// TIA Portal project "dc" (V17)

(* hardware
DEVICE "S7-1200 station_1"  S7-1200 Station
   slot 0: "Rack_0"  S7-1200 Rack  Rack  V1.0
   slot 1: "PLC_1"  CPU 1214C DC/DC/DC  6ES7 214-1AG40-0XB0  V4.4
*)

// ===== PLC "PLC_1"  CPU 1214C DC/DC/DC =====

VAR_GLOBAL   // PLC tag table "Default tag table"
   "Trục Y_Pulse" AT %Q0.2 : Bool;
   "Trục Y_Direction" AT %Q0.3 : Bool;
   "xymove" AT %M110.0 : Bool;
   "xy done" AT %M110.1 : Bool;
   "TRUC_Z_Pulse" AT %Q0.4 : Bool;
   "TRUC_Z_Direction" AT %Q0.5 : Bool;
   "START" AT %I0.0 : Bool;
   "STOP" AT %I0.1 : Bool;
   "E-STOP" AT %I0.2 : Bool;
   "XYZ_home_done" AT %M120.4 : Bool;
   "HMI_X_ActualPos" AT %MD140 : Real;
   "HMI_Y_ActualPos" AT %MD144 : Real;
   "HMI_Z_ActualPos" AT %MD148 : Real;
   "Tag_1" AT %M0.0 : Bool;
   "Tag_2" AT %Q1.0 : Bool;
   "Tag_3" AT %Q1.1 : Bool;
   "Tag_4" AT %M0.1 : Bool;
END_VAR

VAR_GLOBAL   // PLC tag table "TRỤC X"
   "XTrục_Pulse" AT %Q0.0 : Bool;
   "XTrục_Direction" AT %Q0.1 : Bool;
   "X_Enable" AT %M50.0 : Bool;
   "X_Reset" AT %M50.1 : Bool;
   "Jog X+" AT %M50.2 : Bool;
   "Jog X-" AT %M50.3 : Bool;
   "X_Home" AT %M50.4 : Bool;
   "X_MoveAbs" AT %M50.5 : Bool;
   "X_Power_Status" AT %M50.6 : Bool;
   "X_Power_Error" AT %M50.7 : Bool;
   "X_Home_Done" AT %M51.0 : Bool;
   "X_Home_Error" AT %M51.1 : Bool;
   "X_Move_Done" AT %M51.2 : Bool;
   "X_Move_Error" AT %M51.3 : Bool;
   "X_Jog_Error" AT %M51.4 : Bool;
   "X_JogVelocity" AT %MD52 : Real;
   "X_Position" AT %MD56 : Real;
   "X_MoveVelocity" AT %MD60 : Real;
   "X_Home_Sensor" AT %I0.3 : Bool;
   "X_Reset_Done" AT %M51.5 : Bool;
   "X_Reset_Error" AT %M51.6 : Bool;
   "X_Limit_phải" AT %I0.6 : Bool;
   "X_Limit_trái" AT %I0.7 : Bool;
END_VAR

VAR_GLOBAL   // PLC tag table "TRỤC Y"
   "Y_Enable" AT %M70.0 : Bool;
   "Y_Reset" AT %M70.1 : Bool;
   "Jog Y+" AT %M70.2 : Bool;
   "Jog Y-" AT %M70.3 : Bool;
   "Y_Home" AT %M70.4 : Bool;
   "Y_MoveAbs" AT %M70.5 : Bool;
   "Y_Power_Status" AT %M70.6 : Bool;
   "Y_Power_Error" AT %M70.7 : Bool;
   "Y_Home_Done" AT %M71.0 : Bool;
   "Y_Home_Error" AT %M71.1 : Bool;
   "Y_Move_Done" AT %M71.2 : Bool;
   "Y_Move_Error" AT %M71.3 : Bool;
   "Y_Jog_Error" AT %M71.4 : Bool;
   "Y_JogVelocity" AT %MD72 : Real;
   "Y_Position" AT %MD76 : Real;
   "Y_MoveVelocity" AT %MD80 : Real;
   "Y_Home_Sensor" AT %I0.4 : Bool;
   "Y_Reset_Done" AT %M71.5 : Bool;
   "Y_Reset_Error" AT %M71.6 : Bool;
   "Y_Limit_trong" AT %I1.0 : Bool;
   "Y_Limit_ngoai" AT %I1.1 : Bool;
END_VAR

VAR_GLOBAL   // PLC tag table "TRỤC Z"
   "Z_Enable" AT %M90.0 : Bool;
   "Z_Reset" AT %M90.1 : Bool;
   "Jog Z+" AT %M90.2 : Bool;
   "Jog Z-" AT %M90.3 : Bool;
   "Z_Home" AT %M90.4 : Bool;
   "Z_MoveAbs" AT %M90.5 : Bool;
   "Z_Power_Status" AT %M90.6 : Bool;
   "Z_Power_Error" AT %M90.7 : Bool;
   "Z_Home_Done" AT %M91.0 : Bool;
   "Z_Home_Error" AT %M91.1 : Bool;
   "Z_Move_Done" AT %M91.2 : Bool;
   "Z_Move_Error" AT %M91.3 : Bool;
   "Z_Jog_Error" AT %M91.4 : Bool;
   "Z_JogVelocity" AT %MD92 : Real;
   "Z_Position" AT %MD96 : Real;
   "Z_MoveVelocity" AT %MD100 : Real;
   "Z_Home_Sensor" AT %I0.5 : Bool;
   "Z_Reset_Done" AT %M91.5 : Bool;
   "Z_Reset_Error" AT %M91.6 : Bool;
   "Z_Limit_tren" AT %I1.2 : Bool;
   "Z_Limit_duoi" AT %I1.3 : Bool;
END_VAR

VAR_GLOBAL   // PLC tag table "AUTO"
   "HMI_Start" AT %M121.0 : Bool;
   "HMI_Stop" AT %M121.1 : Bool;
   "Start_Cmd" AT %M121.2 : Bool;
   "Stop_Cmd" AT %M121.3 : Bool;
   "AUTO" AT %M120.2 : Bool;
   "AUTO_Step" AT %MW124 : Int;
END_VAR

VAR_GLOBAL   // PLC tag table "Manual"
   "HMI_Manual" AT %M130.0 : Bool;
   "HMI_Auto" AT %M130.1 : Bool;
   "Manual_Mode" AT %M130.2 : Bool;
   "Auto_Mode" AT %M130.3 : Bool;
   "Manual_Ready" AT %M130.4 : Bool;
   "HMI_X_Jog+" AT %M132.0 : Bool;
   "HMI_X_Jog--" AT %M132.1 : Bool;
   "HMI_X_Home" AT %M132.2 : Bool;
   "HMI_X_Reset" AT %M132.3 : Bool;
   "HMI_X_MoveAbs" AT %M132.4 : Bool;
   "HMI_Y_Jog+" AT %M132.5 : Bool;
   "HMI_Y_Jog--" AT %M132.6 : Bool;
   "HMI_Y_Home" AT %M132.7 : Bool;
   "HMI_Y_Reset" AT %M133.0 : Bool;
   "HMI_Y_MoveAbs" AT %M133.1 : Bool;
   "HMI_Z_Jog+" AT %M133.2 : Bool;
   "HMI_Z_Jog-" AT %M133.3 : Bool;
   "HMI_Z_Home" AT %M133.4 : Bool;
   "HMI_Z_Reset" AT %M133.5 : Bool;
   "HMI_Z_MoveAbs" AT %M133.6 : Bool;
END_VAR

DATA_BLOCK "TRUC_X"   // DB1, Motion_DB
{ S7_Optimized_Access := 'TRUE' }
AUTHOR : SIMATIC
FAMILY : BasicMC
NAME : TO_PosAx
VERSION : 7.0
// stored: InstanceOfName TO_PositioningAxis
"TO_PositioningAxis"
BEGIN
   // Axis.PositionLimitsMax_AddressCU = %I0.6
   // Axis.PositionLimitsMin_AddressCU = %I0.7
   // Axis.HomingReferencePointSwitch_AddressCU = %I0.3
   // Axis.LengthUnitNormalized.Distance = 1013
   // Axis.DirectionOutputEnabledCU = TRUE
   // Axis.OnlinePtoModeCU = 16#0000_0002
   // Axis.SelectedChannel2EnumCU = %Q0.1
   // Axis.SelectedChannel1EnumCU = %Q0.0
   // Pulse.MinDeltaDeltaFrequencyCU = 0.004
   // Pulse.MaxDeltaDeltaFrequencyCU = 1.0E+10
   // Pulse.MinDeltaFrequencyCU = 0.005
   // Pulse.MaxDeltaFrequencyCU = 9.5E+9
   // Pulse.MinFrequencyCU = 1.0
   // Pulse.MaxFrequencyCU = 100000.0
   // Pulse.OutputSourceCU = 16#0000_0000
   // Axis.SelectPTO = 0
END_DATA_BLOCK

DATA_BLOCK "Trục Y"   // DB7, Motion_DB
{ S7_Optimized_Access := 'TRUE' }
AUTHOR : SIMATIC
FAMILY : BasicMC
NAME : TO_PosAx
VERSION : 7.0
// stored: InstanceOfName TO_PositioningAxis
"TO_PositioningAxis"
BEGIN
   // Axis.PositionLimitsMax_AddressCU = %I1.1
   // Axis.PositionLimitsMin_AddressCU = %I1.0
   // Axis.HomingReferencePointSwitch_AddressCU = %I0.4
   // Axis.LengthUnitNormalized.Distance = 1013
   // Axis.DirectionOutputEnabledCU = TRUE
   // Axis.OnlinePtoModeCU = 16#0000_0002
   // Axis.SelectedChannel2EnumCU = %Q0.3
   // Axis.SelectedChannel1EnumCU = %Q0.2
   // Pulse.MinDeltaDeltaFrequencyCU = 0.004
   // Pulse.MaxDeltaDeltaFrequencyCU = 1.0E+10
   // Pulse.MinDeltaFrequencyCU = 0.005
   // Pulse.MaxDeltaFrequencyCU = 9.5E+9
   // Pulse.MinFrequencyCU = 1.0
   // Pulse.MaxFrequencyCU = 100000.0
   // Pulse.OutputSourceCU = 16#0000_0000
   // Axis.SelectPTO = 1
   // Axis.OnlinePtoIndexCU = 1
END_DATA_BLOCK

DATA_BLOCK "TRUC_Z"   // DB8, Motion_DB
{ S7_Optimized_Access := 'TRUE' }
AUTHOR : SIMATIC
FAMILY : BasicMC
NAME : TO_PosAx
VERSION : 7.0
// stored: InstanceOfName TO_PositioningAxis
"TO_PositioningAxis"
BEGIN
   // Axis.PositionLimitsMax_AddressCU = %I1.3
   // Axis.PositionLimitsMin_AddressCU = %I1.2
   // Axis.HomingReferencePointSwitch_AddressCU = %I0.5
   // Axis.DirectionOutputEnabledCU = TRUE
   // Axis.LengthUnitNormalized.Distance = 1013
   // Axis.OnlinePtoModeCU = 16#0000_0002
   // Axis.SelectedChannel2EnumCU = %Q0.5
   // Axis.SelectedChannel1EnumCU = %Q0.4
   // Pulse.MinDeltaDeltaFrequencyCU = 0.004
   // Pulse.MaxDeltaDeltaFrequencyCU = 1.0E+10
   // Pulse.MinDeltaFrequencyCU = 0.005
   // Pulse.MaxDeltaFrequencyCU = 9.5E+9
   // Pulse.MinFrequencyCU = 1.0
   // Pulse.MaxFrequencyCU = 30000.0
   // Pulse.OutputSourceCU = 16#0000_0000
   // Axis.SelectPTO = 2
   // Axis.OnlinePtoIndexCU = 2
END_DATA_BLOCK

ORGANIZATION_BLOCK "Main"   // OB1, LAD, ProgramCycle
TITLE = "Main Program Sweep (Cycle)"
{ S7_Optimized_Access := 'TRUE' }
VERSION : 0.1
   VAR_INPUT
      Initial_Call : Bool;   // Initial call of this OB
      Remanence : Bool;   // =True, if remanent data are available
   END_VAR
   VAR_TEMP   // added for the SCL form of the ladder/FBD networks
      _w1 : Bool;
   END_VAR
BEGIN

REGION Network 1
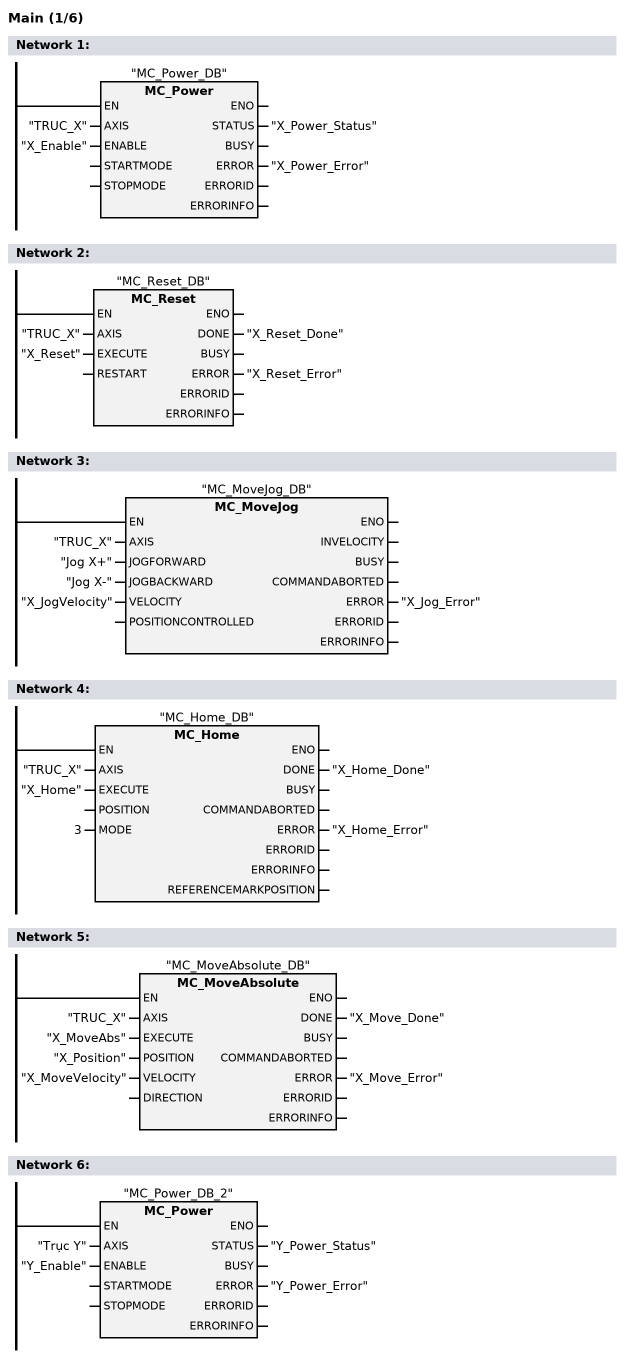
   "MC_Power_DB"(Axis := "TRUC_X", Enable := "X_Enable", Status => "X_Power_Status", Error => "X_Power_Error");   // MC_Power
END_REGION

REGION Network 2
   "MC_Reset_DB"(Axis := "TRUC_X", Execute := "X_Reset", Done => "X_Reset_Done", Error => "X_Reset_Error");   // MC_Reset
END_REGION

REGION Network 3
   "MC_MoveJog_DB"(Axis := "TRUC_X",   // MC_MoveJog
                   JogForward := "Jog X+",
                   JogBackward := "Jog X-",
                   Velocity := "X_JogVelocity",
                   Error => "X_Jog_Error");
END_REGION

REGION Network 4
   "MC_Home_DB"(Axis := "TRUC_X",   // MC_Home
                Execute := "X_Home",
                Mode := 3,
                Done => "X_Home_Done",
                Error => "X_Home_Error");
END_REGION

REGION Network 5
   "MC_MoveAbsolute_DB"(Axis := "TRUC_X",   // MC_MoveAbsolute
                        Execute := "X_MoveAbs",
                        Position := "X_Position",
                        Velocity := "X_MoveVelocity",
                        Done => "X_Move_Done",
                        Error => "X_Move_Error");
END_REGION

REGION Network 6
   "MC_Power_DB_2"(Axis := "Trục Y", Enable := "Y_Enable", Status => "Y_Power_Status", Error => "Y_Power_Error");   // MC_Power
END_REGION

REGION Network 7
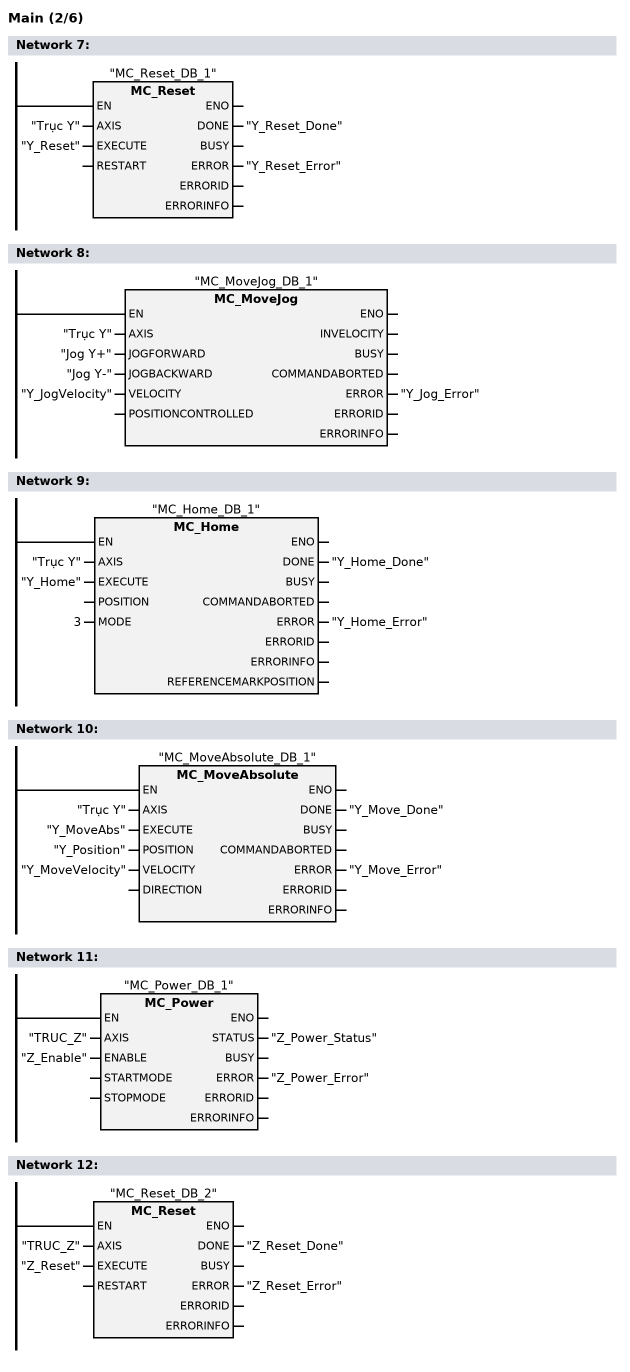
   "MC_Reset_DB_1"(Axis := "Trục Y", Execute := "Y_Reset", Done => "Y_Reset_Done", Error => "Y_Reset_Error");   // MC_Reset
END_REGION

REGION Network 8
   "MC_MoveJog_DB_1"(Axis := "Trục Y",   // MC_MoveJog
                     JogForward := "Jog Y+",
                     JogBackward := "Jog Y-",
                     Velocity := "Y_JogVelocity",
                     Error => "Y_Jog_Error");
END_REGION

REGION Network 9
   "MC_Home_DB_1"(Axis := "Trục Y",   // MC_Home
                  Execute := "Y_Home",
                  Mode := 3,
                  Done => "Y_Home_Done",
                  Error => "Y_Home_Error");
END_REGION

REGION Network 10
   "MC_MoveAbsolute_DB_1"(Axis := "Trục Y",   // MC_MoveAbsolute
                          Execute := "Y_MoveAbs",
                          Position := "Y_Position",
                          Velocity := "Y_MoveVelocity",
                          Done => "Y_Move_Done",
                          Error => "Y_Move_Error");
END_REGION

REGION Network 11
   "MC_Power_DB_1"(Axis := "TRUC_Z", Enable := "Z_Enable", Status => "Z_Power_Status", Error => "Z_Power_Error");   // MC_Power
END_REGION

REGION Network 12
   "MC_Reset_DB_2"(Axis := "TRUC_Z", Execute := "Z_Reset", Done => "Z_Reset_Done", Error => "Z_Reset_Error");   // MC_Reset
END_REGION

REGION Network 13
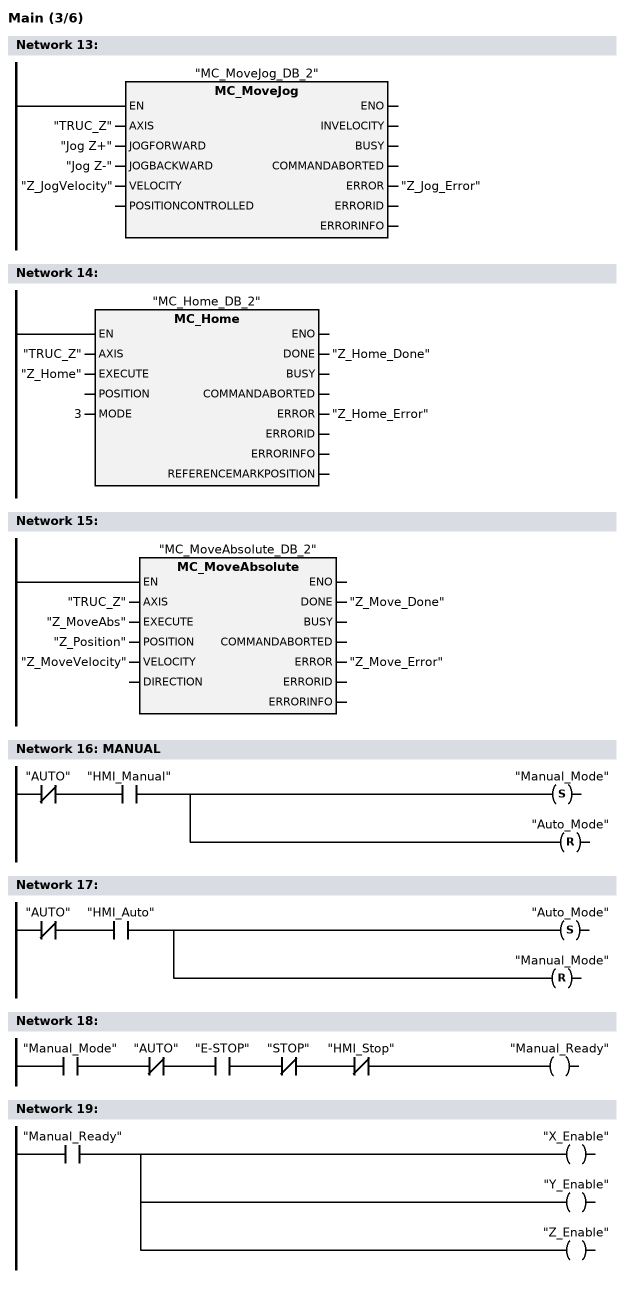
   "MC_MoveJog_DB_2"(Axis := "TRUC_Z",   // MC_MoveJog
                     JogForward := "Jog Z+",
                     JogBackward := "Jog Z-",
                     Velocity := "Z_JogVelocity",
                     Error => "Z_Jog_Error");
END_REGION

REGION Network 14
   "MC_Home_DB_2"(Axis := "TRUC_Z",   // MC_Home
                  Execute := "Z_Home",
                  Mode := 3,
                  Done => "Z_Home_Done",
                  Error => "Z_Home_Error");
END_REGION

REGION Network 15
   "MC_MoveAbsolute_DB_2"(Axis := "TRUC_Z",   // MC_MoveAbsolute
                          Execute := "Z_MoveAbs",
                          Position := "Z_Position",
                          Velocity := "Z_MoveVelocity",
                          Done => "Z_Move_Done",
                          Error => "Z_Move_Error");
END_REGION

REGION Network 16: MANUAL
   RUNG wire#powerrail
      I_Contact( "AUTO" )
      Contact( "HMI_Manual" )
      wire#w1
      S_Coil( "Manual_Mode" )
   END_RUNG
   RUNG wire#w1
      R_Coil( "Auto_Mode" )
   END_RUNG
   // the same network as SCL:
   IF NOT "AUTO" AND "HMI_Manual" THEN
       "Manual_Mode" := TRUE;
       "Auto_Mode" := FALSE;
   END_IF;
END_REGION

REGION Network 17
   RUNG wire#powerrail
      I_Contact( "AUTO" )
      Contact( "HMI_Auto" )
      wire#w1
      S_Coil( "Auto_Mode" )
   END_RUNG
   RUNG wire#w1
      R_Coil( "Manual_Mode" )
   END_RUNG
   // the same network as SCL:
   IF NOT "AUTO" AND "HMI_Auto" THEN
       "Auto_Mode" := TRUE;
       "Manual_Mode" := FALSE;
   END_IF;
END_REGION

REGION Network 18
   RUNG wire#powerrail
      Contact( "Manual_Mode" )
      I_Contact( "AUTO" )
      Contact( "E-STOP" )
      I_Contact( "STOP" )
      I_Contact( "HMI_Stop" )
      Coil( "Manual_Ready" )
   END_RUNG
   // the same network as SCL:
   "Manual_Ready" := "Manual_Mode" AND NOT "AUTO" AND "E-STOP" AND NOT "STOP" AND NOT "HMI_Stop";
END_REGION

REGION Network 19
   RUNG wire#powerrail
      Contact( "Manual_Ready" )
      wire#w1
      Coil( "X_Enable" )
   END_RUNG
   RUNG wire#w1
      Coil( "Y_Enable" )
   END_RUNG
   RUNG wire#w1
      Coil( "Z_Enable" )
   END_RUNG
   // the same network as SCL:
   "X_Enable" := "Manual_Ready";
   "Y_Enable" := "Manual_Ready";
   "Z_Enable" := "Manual_Ready";
END_REGION

REGION Network 20
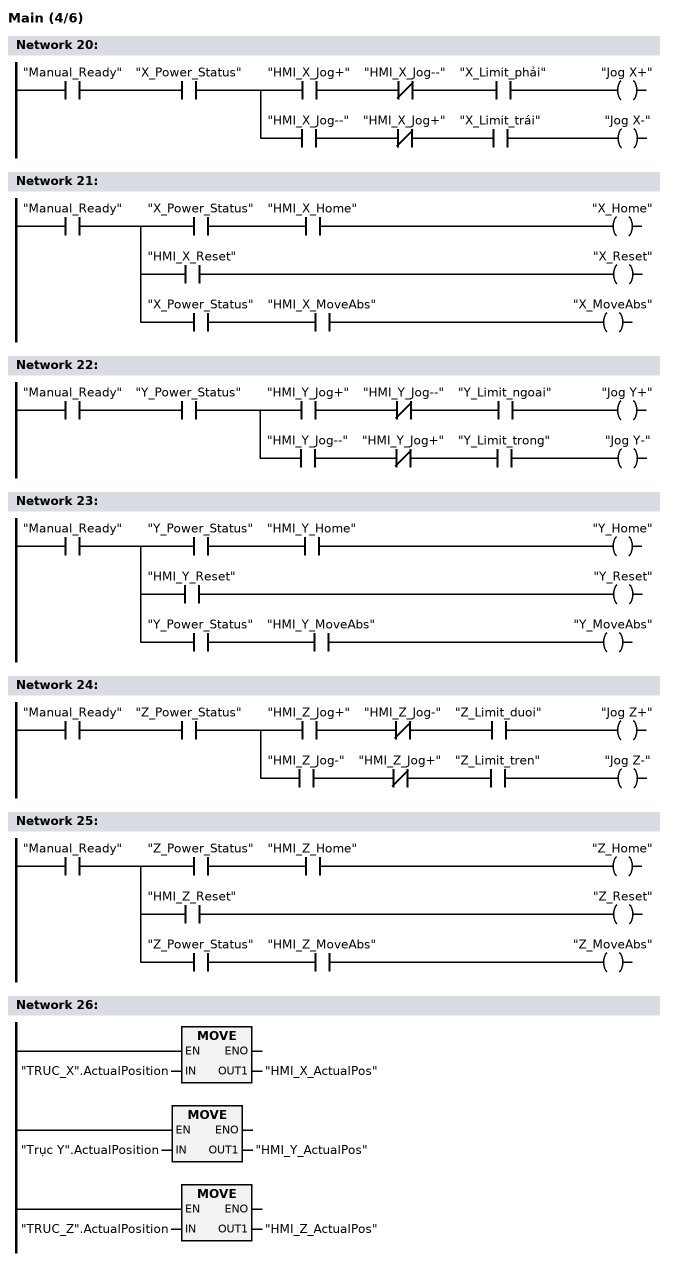
   RUNG wire#powerrail
      Contact( "Manual_Ready" )
      Contact( "X_Power_Status" )
      wire#w1
      Contact( "HMI_X_Jog+" )
      I_Contact( "HMI_X_Jog--" )
      Contact( "X_Limit_phải" )
      Coil( "Jog X+" )
   END_RUNG
   RUNG wire#w1
      Contact( "HMI_X_Jog--" )
      I_Contact( "HMI_X_Jog+" )
      Contact( "X_Limit_trái" )
      Coil( "Jog X-" )
   END_RUNG
   // the same network as SCL:
   #_w1 := "Manual_Ready" AND "X_Power_Status";
   "Jog X+" := #_w1 AND "HMI_X_Jog+" AND NOT "HMI_X_Jog--" AND "X_Limit_phải";
   "Jog X-" := #_w1 AND "HMI_X_Jog--" AND NOT "HMI_X_Jog+" AND "X_Limit_trái";
END_REGION

REGION Network 21
   RUNG wire#powerrail
      Contact( "Manual_Ready" )
      wire#w1
      Contact( "X_Power_Status" )
      Contact( "HMI_X_Home" )
      Coil( "X_Home" )
   END_RUNG
   RUNG wire#w1
      Contact( "HMI_X_Reset" )
      Coil( "X_Reset" )
   END_RUNG
   RUNG wire#w1
      Contact( "X_Power_Status" )
      Contact( "HMI_X_MoveAbs" )
      Coil( "X_MoveAbs" )
   END_RUNG
   // the same network as SCL:
   "X_Home" := "Manual_Ready" AND "X_Power_Status" AND "HMI_X_Home";
   "X_Reset" := "Manual_Ready" AND "HMI_X_Reset";
   "X_MoveAbs" := "Manual_Ready" AND "X_Power_Status" AND "HMI_X_MoveAbs";
END_REGION

REGION Network 22
   RUNG wire#powerrail
      Contact( "Manual_Ready" )
      Contact( "Y_Power_Status" )
      wire#w1
      Contact( "HMI_Y_Jog+" )
      I_Contact( "HMI_Y_Jog--" )
      Contact( "Y_Limit_ngoai" )
      Coil( "Jog Y+" )
   END_RUNG
   RUNG wire#w1
      Contact( "HMI_Y_Jog--" )
      I_Contact( "HMI_Y_Jog+" )
      Contact( "Y_Limit_trong" )
      Coil( "Jog Y-" )
   END_RUNG
   // the same network as SCL:
   #_w1 := "Manual_Ready" AND "Y_Power_Status";
   "Jog Y+" := #_w1 AND "HMI_Y_Jog+" AND NOT "HMI_Y_Jog--" AND "Y_Limit_ngoai";
   "Jog Y-" := #_w1 AND "HMI_Y_Jog--" AND NOT "HMI_Y_Jog+" AND "Y_Limit_trong";
END_REGION

REGION Network 23
   RUNG wire#powerrail
      Contact( "Manual_Ready" )
      wire#w1
      Contact( "Y_Power_Status" )
      Contact( "HMI_Y_Home" )
      Coil( "Y_Home" )
   END_RUNG
   RUNG wire#w1
      Contact( "HMI_Y_Reset" )
      Coil( "Y_Reset" )
   END_RUNG
   RUNG wire#w1
      Contact( "Y_Power_Status" )
      Contact( "HMI_Y_MoveAbs" )
      Coil( "Y_MoveAbs" )
   END_RUNG
   // the same network as SCL:
   "Y_Home" := "Manual_Ready" AND "Y_Power_Status" AND "HMI_Y_Home";
   "Y_Reset" := "Manual_Ready" AND "HMI_Y_Reset";
   "Y_MoveAbs" := "Manual_Ready" AND "Y_Power_Status" AND "HMI_Y_MoveAbs";
END_REGION

REGION Network 24
   RUNG wire#powerrail
      Contact( "Manual_Ready" )
      Contact( "Z_Power_Status" )
      wire#w1
      Contact( "HMI_Z_Jog+" )
      I_Contact( "HMI_Z_Jog-" )
      Contact( "Z_Limit_duoi" )
      Coil( "Jog Z+" )
   END_RUNG
   RUNG wire#w1
      Contact( "HMI_Z_Jog-" )
      I_Contact( "HMI_Z_Jog+" )
      Contact( "Z_Limit_tren" )
      Coil( "Jog Z-" )
   END_RUNG
   // the same network as SCL:
   #_w1 := "Manual_Ready" AND "Z_Power_Status";
   "Jog Z+" := #_w1 AND "HMI_Z_Jog+" AND NOT "HMI_Z_Jog-" AND "Z_Limit_duoi";
   "Jog Z-" := #_w1 AND "HMI_Z_Jog-" AND NOT "HMI_Z_Jog+" AND "Z_Limit_tren";
END_REGION

REGION Network 25
   RUNG wire#powerrail
      Contact( "Manual_Ready" )
      wire#w1
      Contact( "Z_Power_Status" )
      Contact( "HMI_Z_Home" )
      Coil( "Z_Home" )
   END_RUNG
   RUNG wire#w1
      Contact( "HMI_Z_Reset" )
      Coil( "Z_Reset" )
   END_RUNG
   RUNG wire#w1
      Contact( "Z_Power_Status" )
      Contact( "HMI_Z_MoveAbs" )
      Coil( "Z_MoveAbs" )
   END_RUNG
   // the same network as SCL:
   "Z_Home" := "Manual_Ready" AND "Z_Power_Status" AND "HMI_Z_Home";
   "Z_Reset" := "Manual_Ready" AND "HMI_Z_Reset";
   "Z_MoveAbs" := "Manual_Ready" AND "Z_Power_Status" AND "HMI_Z_MoveAbs";
END_REGION

REGION Network 26
   RUNG wire#powerrail
      Move(in := "TRUC_X".ActualPosition, out1 => "HMI_X_ActualPos")
   END_RUNG
   RUNG wire#powerrail
      Move(in := "Trục Y".ActualPosition, out1 => "HMI_Y_ActualPos")
   END_RUNG
   RUNG wire#powerrail
      Move(in := "TRUC_Z".ActualPosition, out1 => "HMI_Z_ActualPos")
   END_RUNG
   // the same network as SCL:
   "HMI_X_ActualPos" := "TRUC_X".ActualPosition;
   "HMI_Y_ActualPos" := "Trục Y".ActualPosition;
   "HMI_Z_ActualPos" := "TRUC_Z".ActualPosition;
END_REGION

REGION Network 27
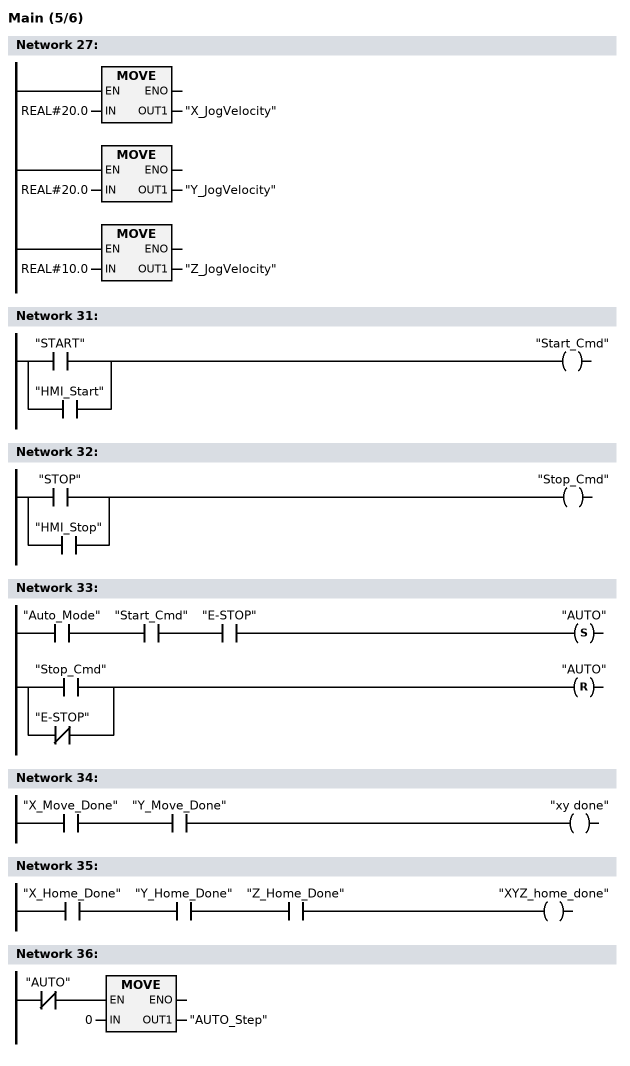
   RUNG wire#powerrail
      Move(in := REAL#20.0, out1 => "X_JogVelocity")
   END_RUNG
   RUNG wire#powerrail
      Move(in := REAL#20.0, out1 => "Y_JogVelocity")
   END_RUNG
   RUNG wire#powerrail
      Move(in := REAL#10.0, out1 => "Z_JogVelocity")
   END_RUNG
   // the same network as SCL:
   "X_JogVelocity" := REAL#20.0;
   "Y_JogVelocity" := REAL#20.0;
   "Z_JogVelocity" := REAL#10.0;
END_REGION

REGION Network 31
   RUNG wire#powerrail
      Contact( "START" )
      wire#w1
      Coil( "Start_Cmd" )
   END_RUNG
   RUNG wire#powerrail
      Contact( "HMI_Start" )
   END_RUNG wire#w1
   // the same network as SCL:
   "Start_Cmd" := "START" OR "HMI_Start";
END_REGION

REGION Network 32
   RUNG wire#powerrail
      Contact( "STOP" )
      wire#w1
      Coil( "Stop_Cmd" )
   END_RUNG
   RUNG wire#powerrail
      Contact( "HMI_Stop" )
   END_RUNG wire#w1
   // the same network as SCL:
   "Stop_Cmd" := "STOP" OR "HMI_Stop";
END_REGION

REGION Network 33
   RUNG wire#powerrail
      Contact( "Auto_Mode" )
      Contact( "Start_Cmd" )
      Contact( "E-STOP" )
      S_Coil( "AUTO" )
   END_RUNG
   RUNG wire#powerrail
      Contact( "Stop_Cmd" )
      wire#w1
      R_Coil( "AUTO" )
   END_RUNG
   RUNG wire#powerrail
      I_Contact( "E-STOP" )
   END_RUNG wire#w1
   // the same network as SCL:
   IF "Auto_Mode" AND "Start_Cmd" AND "E-STOP" THEN "AUTO" := TRUE; END_IF;
   IF "Stop_Cmd" OR NOT "E-STOP" THEN "AUTO" := FALSE; END_IF;
END_REGION

REGION Network 34
   RUNG wire#powerrail
      Contact( "X_Move_Done" )
      Contact( "Y_Move_Done" )
      Coil( "xy done" )
   END_RUNG
   // the same network as SCL:
   "xy done" := "X_Move_Done" AND "Y_Move_Done";
END_REGION

REGION Network 35
   RUNG wire#powerrail
      Contact( "X_Home_Done" )
      Contact( "Y_Home_Done" )
      Contact( "Z_Home_Done" )
      Coil( "XYZ_home_done" )
   END_RUNG
   // the same network as SCL:
   "XYZ_home_done" := "X_Home_Done" AND "Y_Home_Done" AND "Z_Home_Done";
END_REGION

REGION Network 36
   RUNG wire#powerrail
      I_Contact( "AUTO" )
      Move(in := 0, out1 => "AUTO_Step")
   END_RUNG
   // the same network as SCL:
   IF NOT "AUTO" THEN "AUTO_Step" := 0; END_IF;
END_REGION

REGION Network 37
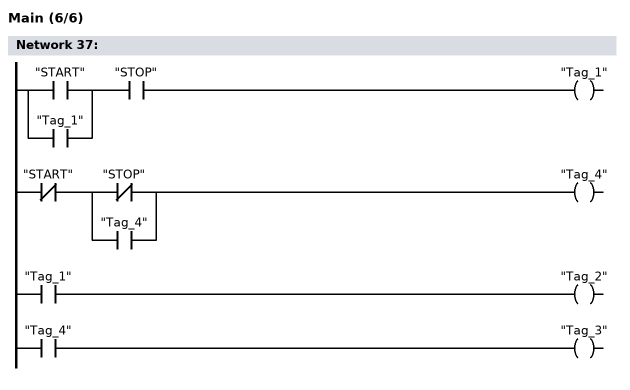
   RUNG wire#powerrail
      Contact( "START" )
      wire#w1
      Contact( "STOP" )
      Coil( "Tag_1" )
   END_RUNG
   RUNG wire#powerrail
      Contact( "Tag_1" )
   END_RUNG wire#w1
   RUNG wire#powerrail
      I_Contact( "START" )
      wire#w2
      I_Contact( "STOP" )
      wire#w3
      Coil( "Tag_4" )
   END_RUNG
   RUNG wire#w2
      Contact( "Tag_4" )
   END_RUNG wire#w3
   RUNG wire#powerrail
      Contact( "Tag_1" )
      Coil( "Tag_2" )
   END_RUNG
   RUNG wire#powerrail
      Contact( "Tag_4" )
      Coil( "Tag_3" )
   END_RUNG
   // the same network as SCL:
   "Tag_1" := ("START" OR "Tag_1") AND "STOP";
   "Tag_4" := NOT "START" AND (NOT "STOP" OR "Tag_4");
   "Tag_2" := "Tag_1";
   "Tag_3" := "Tag_4";
END_REGION
END_ORGANIZATION_BLOCK